(* IEC 61131-3 sources: plc-st-coding-agent/progress/evidence/f14_v11_public_20261113/jobs/custom_deepseek-v4pro (part 2) *)

(* ---- public-hard-02.candidate_03.st ---- *)
TYPE ProcessControl_State : (PC_IDLE, PC_MOVING, PC_WAITING); END_TYPE;

FUNCTION_BLOCK FlexibleProcessingControl
VAR_INPUT
    processLength : USINT;
    sensor1 : BOOL;
    sensor2 : BOOL;
    sensor3 : BOOL;
    sensor4 : BOOL;
    sensor5 : BOOL;
    station1Start : BOOL;
    station2Complete : BOOL;
    station3Complete : BOOL;
    station4Complete : BOOL;
    processSequence : ARRAY[1..8] OF USINT;
END_VAR
VAR_OUTPUT
    conveyorLeft : BOOL;
    conveyorRight : BOOL;
END_VAR
VAR
    state : ProcessControl_State := PC_IDLE;
    currentStation : USINT := 1;
    currentIndex : USINT := 1;
    targetStation : USINT := 0;
    targetSensor : BOOL := FALSE;
    local_rt_start : R_TRIG;
    local_rt_st2 : R_TRIG;
    local_rt_st3 : R_TRIG;
    local_rt_st4 : R_TRIG;
END_VAR

(*
ENGINEERING_CONTRACT
  conveyorLeft / conveyorRight activation: PC_MOVING state and target direction >/< currentStation (PUB001-PUB002).
  Retention/hold: outputs stay on each scan while PC_MOVING until target sensor TRUE (PUB002).
  Explicit reset/deactivation: sensor at target station stops motion and sets both outputs FALSE; next start new product.
  Same-scan priority: start request processed only in PC_IDLE; arrival stop and completion advancement are mutually exclusive by state.
  Units/boundaries: processLength 1..8; processSequence index 1..8; currentStation 1..5; final active entry 5 (PUB003).
  Direction: target > current -> conveyorRight; target < current -> conveyorLeft; target == current -> no movement, treated as arrived.
  Completion edge: rising edge of station2Complete/3/4Complete triggers next step.
  Unspecified: equal consecutive station entries skip movement and wait for completion; simultaneous completion inputs while WAITING use current station only.
*)

(* CONTRACT_RULES [] *)

local_rt_start(CLK := station1Start AND sensor1);
local_rt_st2(CLK := station2Complete);
local_rt_st3(CLK := station3Complete);
local_rt_st4(CLK := station4Complete);

CASE state OF
    PC_IDLE:
        conveyorLeft := FALSE;
        conveyorRight := FALSE;
        IF local_rt_start.Q THEN
            currentIndex := 1;
            currentStation := 1;
            targetStation := processSequence[currentIndex];
            IF targetStation = currentStation THEN
                IF targetStation = 5 THEN
                    state := PC_IDLE;
                ELSE
                    state := PC_WAITING;
                END_IF;
            ELSE
                state := PC_MOVING;
            END_IF;
        END_IF;

    PC_MOVING:
        targetSensor := FALSE;
        CASE targetStation OF
            2: targetSensor := sensor2;
            3: targetSensor := sensor3;
            4: targetSensor := sensor4;
            5: targetSensor := sensor5;
        END_CASE;

        IF targetStation > currentStation THEN
            conveyorLeft := FALSE;
            conveyorRight := TRUE;
        ELSIF targetStation < currentStation THEN
            conveyorLeft := TRUE;
            conveyorRight := FALSE;
        ELSE
            conveyorLeft := FALSE;
            conveyorRight := FALSE;
        END_IF;

        IF targetSensor THEN
            conveyorLeft := FALSE;
            conveyorRight := FALSE;
            currentStation := targetStation;
            IF targetStation = 5 THEN
                state := PC_IDLE;
            ELSE
                state := PC_WAITING;
            END_IF;
        END_IF;

    PC_WAITING:
        conveyorLeft := FALSE;
        conveyorRight := FALSE;
        IF (currentStation = 2 AND local_rt_st2.Q) OR
           (currentStation = 3 AND local_rt_st3.Q) OR
           (currentStation = 4 AND local_rt_st4.Q) THEN
            IF currentIndex < processLength THEN
                currentIndex := currentIndex + 1;
                targetStation := processSequence[currentIndex];
                IF targetStation = currentStation THEN
                    IF targetStation = 5 THEN
                        state := PC_IDLE;
                    ELSE
                        state := PC_WAITING;
                    END_IF;
                ELSE
                    state := PC_MOVING;
                END_IF;
            ELSE
                state := PC_IDLE;
            END_IF;
        END_IF;
END_CASE;

(* Same-scan output update after any state transition *)
IF state = PC_MOVING THEN
    IF targetStation > currentStation THEN
        conveyorLeft := FALSE;
        conveyorRight := TRUE;
    ELSIF targetStation < currentStation THEN
        conveyorLeft := TRUE;
        conveyorRight := FALSE;
    ELSE
        conveyorLeft := FALSE;
        conveyorRight := FALSE;
    END_IF;
ELSE
    conveyorLeft := FALSE;
    conveyorRight := FALSE;
END_IF;

END_FUNCTION_BLOCK

(* ---- public-hard-02.candidate_04.st ---- *)
TYPE ProcessControl_State : (PC_IDLE, PC_MOVING, PC_WAITING); END_TYPE;

FUNCTION_BLOCK FlexibleProcessingControl
VAR_INPUT
    processLength : USINT;
    sensor1 : BOOL;
    sensor2 : BOOL;
    sensor3 : BOOL;
    sensor4 : BOOL;
    sensor5 : BOOL;
    station1Start : BOOL;
    station2Complete : BOOL;
    station3Complete : BOOL;
    station4Complete : BOOL;
    processSequence : ARRAY[1..8] OF USINT;
END_VAR
VAR_OUTPUT
    conveyorLeft : BOOL;
    conveyorRight : BOOL;
END_VAR
VAR
    state : ProcessControl_State := PC_IDLE;
    currentStation : USINT := 1;
    currentIndex : USINT := 1;
    targetStation : USINT := 0;
    targetSensor : BOOL := FALSE;
    local_rt_start : R_TRIG;
    local_rt_st2 : R_TRIG;
    local_rt_st3 : R_TRIG;
    local_rt_st4 : R_TRIG;
END_VAR

(*
ENGINEERING_CONTRACT
  conveyorLeft / conveyorRight activation: PC_MOVING state and target direction >/< currentStation (PUB001-PUB002).
  Retention/hold: outputs stay on each scan while PC_MOVING until target sensor TRUE (PUB002).
  Explicit reset/deactivation: sensor at target station stops motion and sets both outputs FALSE; next start new product.
  Same-scan priority: start request processed only in PC_IDLE; arrival stop and completion advancement are mutually exclusive by state.
  Units/boundaries: processLength 1..8; processSequence index 1..8; currentStation 1..5; final active entry 5 (PUB003).
  Direction: target > current -> conveyorRight; target < current -> conveyorLeft; target == current -> no movement, treated as arrived.
  Completion edge: rising edge of station2Complete/3/4Complete triggers next step.
  Unspecified: equal consecutive station entries skip movement and wait for completion; simultaneous completion inputs while WAITING use current station only.
  Same-scan start with target sensor already active causes immediate arrival handling without starting conveyor.
*)

(* CONTRACT_RULES [] *)

local_rt_start(CLK := station1Start AND sensor1);
local_rt_st2(CLK := station2Complete);
local_rt_st3(CLK := station3Complete);
local_rt_st4(CLK := station4Complete);

CASE state OF
    PC_IDLE:
        conveyorLeft := FALSE;
        conveyorRight := FALSE;
        IF local_rt_start.Q THEN
            currentIndex := 1;
            currentStation := 1;
            targetStation := processSequence[currentIndex];
            IF targetStation = currentStation THEN
                IF targetStation = 5 THEN
                    state := PC_IDLE;
                ELSE
                    state := PC_WAITING;
                END_IF;
            ELSE
                targetSensor := FALSE;
                CASE targetStation OF
                    2: targetSensor := sensor2;
                    3: targetSensor := sensor3;
                    4: targetSensor := sensor4;
                    5: targetSensor := sensor5;
                END_CASE;
                IF targetSensor THEN
                    currentStation := targetStation;
                    IF targetStation = 5 THEN
                        state := PC_IDLE;
                    ELSE
                        state := PC_WAITING;
                    END_IF;
                ELSE
                    state := PC_MOVING;
                END_IF;
            END_IF;
        END_IF;

    PC_MOVING:
        targetSensor := FALSE;
        CASE targetStation OF
            2: targetSensor := sensor2;
            3: targetSensor := sensor3;
            4: targetSensor := sensor4;
            5: targetSensor := sensor5;
        END_CASE;

        IF targetStation > currentStation THEN
            conveyorLeft := FALSE;
            conveyorRight := TRUE;
        ELSIF targetStation < currentStation THEN
            conveyorLeft := TRUE;
            conveyorRight := FALSE;
        ELSE
            conveyorLeft := FALSE;
            conveyorRight := FALSE;
        END_IF;

        IF targetSensor THEN
            conveyorLeft := FALSE;
            conveyorRight := FALSE;
            currentStation := targetStation;
            IF targetStation = 5 THEN
                state := PC_IDLE;
            ELSE
                state := PC_WAITING;
            END_IF;
        END_IF;

    PC_WAITING:
        conveyorLeft := FALSE;
        conveyorRight := FALSE;
        IF (currentStation = 2 AND local_rt_st2.Q) OR
           (currentStation = 3 AND local_rt_st3.Q) OR
           (currentStation = 4 AND local_rt_st4.Q) THEN
            IF currentIndex < processLength THEN
                currentIndex := currentIndex + 1;
                targetStation := processSequence[currentIndex];
                IF targetStation = currentStation THEN
                    IF targetStation = 5 THEN
                        state := PC_IDLE;
                    ELSE
                        state := PC_WAITING;
                    END_IF;
                ELSE
                    state := PC_MOVING;
                END_IF;
            ELSE
                state := PC_IDLE;
            END_IF;
        END_IF;
END_CASE;

(* Same-scan output update after any state transition *)
IF state = PC_MOVING THEN
    IF targetStation > currentStation THEN
        conveyorLeft := FALSE;
        conveyorRight := TRUE;
    ELSIF targetStation < currentStation THEN
        conveyorLeft := TRUE;
        conveyorRight := FALSE;
    ELSE
        conveyorLeft := FALSE;
        conveyorRight := FALSE;
    END_IF;
ELSE
    conveyorLeft := FALSE;
    conveyorRight := FALSE;
END_IF;

END_FUNCTION_BLOCK

(* ---- public-hard-02.raw_candidate_01.st ---- *)
TYPE ProcessControl_State : (PC_IDLE, PC_MOVING, PC_WAITING); END_TYPE

FUNCTION_BLOCK FlexibleProcessingControl
VAR_INPUT
    processLength : USINT;
    sensor1 : BOOL;
    sensor2 : BOOL;
    sensor3 : BOOL;
    sensor4 : BOOL;
    sensor5 : BOOL;
    station1Start : BOOL;
    station2Complete : BOOL;
    station3Complete : BOOL;
    station4Complete : BOOL;
    processSequence : ARRAY[1..8] OF USINT;
END_VAR
VAR_OUTPUT
    conveyorLeft : BOOL;
    conveyorRight : BOOL;
END_VAR
VAR
    state : ProcessControl_State := PC_IDLE;
    currentStation : USINT := 1;
    currentIndex : USINT := 1;
    targetStation : USINT := 0;
    targetSensor : BOOL := FALSE;
    local_rt_start : R_TRIG;
    local_rt_st2 : R_TRIG;
    local_rt_st3 : R_TRIG;
    local_rt_st4 : R_TRIG;
END_VAR

(*
ENGINEERING_CONTRACT
  conveyorLeft / conveyorRight activation: PC_MOVING state and target direction >/< currentStation (PUB001-PUB002).
  Retention/hold: outputs stay on each scan while PC_MOVING until target sensor TRUE (PUB002).
  Explicit reset/deactivation: sensor at target station stops motion and sets both outputs FALSE; next start new product.
  Same-scan priority: start request processed only in PC_IDLE; arrival stop and completion advancement are mutually exclusive by state.
  Units/boundaries: processLength 1..8; processSequence index 1..8; currentStation 1..5; final active entry 5 (PUB003).
  Direction: target > current -> conveyorRight; target < current -> conveyorLeft; target == current -> no movement, treated as arrived.
  Completion edge: rising edge of station2Complete/3/4Complete triggers next step.
  Unspecified: equal consecutive station entries skip movement and wait for completion; simultaneous completion inputs while WAITING use current station only.
*)

(* CONTRACT_RULES [] *)

local_rt_start(CLK := station1Start);
local_rt_st2(CLK := station2Complete);
local_rt_st3(CLK := station3Complete);
local_rt_st4(CLK := station4Complete);

CASE state OF
    PC_IDLE:
        conveyorLeft := FALSE;
        conveyorRight := FALSE;
        IF local_rt_start.Q AND sensor1 THEN
            currentIndex := 1;
            currentStation := 1;
            targetStation := processSequence[currentIndex];
            IF targetStation = currentStation THEN
                IF targetStation = 5 THEN
                    state := PC_IDLE;
                ELSE
                    state := PC_WAITING;
                END_IF;
            ELSE
                state := PC_MOVING;
            END_IF;
        END_IF;

    PC_MOVING:
        targetSensor := FALSE;
        CASE targetStation OF
            2: targetSensor := sensor2;
            3: targetSensor := sensor3;
            4: targetSensor := sensor4;
            5: targetSensor := sensor5;
        END_CASE;

        IF targetStation > currentStation THEN
            conveyorLeft := FALSE;
            conveyorRight := TRUE;
        ELSIF targetStation < currentStation THEN
            conveyorLeft := TRUE;
            conveyorRight := FALSE;
        ELSE
            conveyorLeft := FALSE;
            conveyorRight := FALSE;
        END_IF;

        IF targetSensor THEN
            conveyorLeft := FALSE;
            conveyorRight := FALSE;
            currentStation := targetStation;
            IF targetStation = 5 THEN
                state := PC_IDLE;
            ELSE
                state := PC_WAITING;
            END_IF;
        END_IF;

    PC_WAITING:
        conveyorLeft := FALSE;
        conveyorRight := FALSE;
        IF (currentStation = 2 AND local_rt_st2.Q) OR
           (currentStation = 3 AND local_rt_st3.Q) OR
           (currentStation = 4 AND local_rt_st4.Q) THEN
            IF currentIndex < processLength THEN
                currentIndex := currentIndex + 1;
                targetStation := processSequence[currentIndex];
                IF targetStation = currentStation THEN
                    IF targetStation = 5 THEN
                        state := PC_IDLE;
                    ELSE
                        state := PC_WAITING;
                    END_IF;
                ELSE
                    state := PC_MOVING;
                END_IF;
            ELSE
                state := PC_IDLE;
            END_IF;
        END_IF;
END_CASE;

(* ---- public-hard-02.raw_candidate_02.st ---- *)
TYPE ProcessControl_State : (PC_IDLE, PC_MOVING, PC_WAITING); END_TYPE;

FUNCTION_BLOCK FlexibleProcessingControl
VAR_INPUT
    processLength : USINT;
    sensor1 : BOOL;
    sensor2 : BOOL;
    sensor3 : BOOL;
    sensor4 : BOOL;
    sensor5 : BOOL;
    station1Start : BOOL;
    station2Complete : BOOL;
    station3Complete : BOOL;
    station4Complete : BOOL;
    processSequence : ARRAY[1..8] OF USINT;
END_VAR
VAR_OUTPUT
    conveyorLeft : BOOL;
    conveyorRight : BOOL;
END_VAR
VAR
    state : ProcessControl_State := PC_IDLE;
    currentStation : USINT := 1;
    currentIndex : USINT := 1;
    targetStation : USINT := 0;
    targetSensor : BOOL := FALSE;
    local_rt_start : R_TRIG;
    local_rt_st2 : R_TRIG;
    local_rt_st3 : R_TRIG;
    local_rt_st4 : R_TRIG;
END_VAR

(*
ENGINEERING_CONTRACT
  conveyorLeft / conveyorRight activation: PC_MOVING state and target direction >/< currentStation (PUB001-PUB002).
  Retention/hold: outputs stay on each scan while PC_MOVING until target sensor TRUE (PUB002).
  Explicit reset/deactivation: sensor at target station stops motion and sets both outputs FALSE; next start new product.
  Same-scan priority: start request processed only in PC_IDLE; arrival stop and completion advancement are mutually exclusive by state.
  Units/boundaries: processLength 1..8; processSequence index 1..8; currentStation 1..5; final active entry 5 (PUB003).
  Direction: target > current -> conveyorRight; target < current -> conveyorLeft; target == current -> no movement, treated as arrived.
  Completion edge: rising edge of station2Complete/3/4Complete triggers next step.
  Unspecified: equal consecutive station entries skip movement and wait for completion; simultaneous completion inputs while WAITING use current station only.
*)

(* CONTRACT_RULES [] *)

local_rt_start(CLK := station1Start);
local_rt_st2(CLK := station2Complete);
local_rt_st3(CLK := station3Complete);
local_rt_st4(CLK := station4Complete);

CASE state OF
    PC_IDLE:
        conveyorLeft := FALSE;
        conveyorRight := FALSE;
        IF local_rt_start.Q AND sensor1 THEN
            currentIndex := 1;
            currentStation := 1;
            targetStation := processSequence[currentIndex];
            IF targetStation = currentStation THEN
                IF targetStation = 5 THEN
                    state := PC_IDLE;
                ELSE
                    state := PC_WAITING;
                END_IF;
            ELSE
                state := PC_MOVING;
            END_IF;
        END_IF;

    PC_MOVING:
        targetSensor := FALSE;
        CASE targetStation OF
            2: targetSensor := sensor2;
            3: targetSensor := sensor3;
            4: targetSensor := sensor4;
            5: targetSensor := sensor5;
        END_CASE;

        IF targetStation > currentStation THEN
            conveyorLeft := FALSE;
            conveyorRight := TRUE;
        ELSIF targetStation < currentStation THEN
            conveyorLeft := TRUE;
            conveyorRight := FALSE;
        ELSE
            conveyorLeft := FALSE;
            conveyorRight := FALSE;
        END_IF;

        IF targetSensor THEN
            conveyorLeft := FALSE;
            conveyorRight := FALSE;
            currentStation := targetStation;
            IF targetStation = 5 THEN
                state := PC_IDLE;
            ELSE
                state := PC_WAITING;
            END_IF;
        END_IF;

    PC_WAITING:
        conveyorLeft := FALSE;
        conveyorRight := FALSE;
        IF (currentStation = 2 AND local_rt_st2.Q) OR
           (currentStation = 3 AND local_rt_st3.Q) OR
           (currentStation = 4 AND local_rt_st4.Q) THEN
            IF currentIndex < processLength THEN
                currentIndex := currentIndex + 1;
                targetStation := processSequence[currentIndex];
                IF targetStation = currentStation THEN
                    IF targetStation = 5 THEN
                        state := PC_IDLE;
                    ELSE
                        state := PC_WAITING;
                    END_IF;
                ELSE
                    state := PC_MOVING;
                END_IF;
            ELSE
                state := PC_IDLE;
            END_IF;
        END_IF;
END_CASE;

END_FUNCTION_BLOCK

(* ---- public-hard-02.raw_candidate_03.st ---- *)
TYPE ProcessControl_State : (PC_IDLE, PC_MOVING, PC_WAITING); END_TYPE;

FUNCTION_BLOCK FlexibleProcessingControl
VAR_INPUT
    processLength : USINT;
    sensor1 : BOOL;
    sensor2 : BOOL;
    sensor3 : BOOL;
    sensor4 : BOOL;
    sensor5 : BOOL;
    station1Start : BOOL;
    station2Complete : BOOL;
    station3Complete : BOOL;
    station4Complete : BOOL;
    processSequence : ARRAY[1..8] OF USINT;
END_VAR
VAR_OUTPUT
    conveyorLeft : BOOL;
    conveyorRight : BOOL;
END_VAR
VAR
    state : ProcessControl_State := PC_IDLE;
    currentStation : USINT := 1;
    currentIndex : USINT := 1;
    targetStation : USINT := 0;
    targetSensor : BOOL := FALSE;
    local_rt_start : R_TRIG;
    local_rt_st2 : R_TRIG;
    local_rt_st3 : R_TRIG;
    local_rt_st4 : R_TRIG;
END_VAR

(*
ENGINEERING_CONTRACT
  conveyorLeft / conveyorRight activation: PC_MOVING state and target direction >/< currentStation (PUB001-PUB002).
  Retention/hold: outputs stay on each scan while PC_MOVING until target sensor TRUE (PUB002).
  Explicit reset/deactivation: sensor at target station stops motion and sets both outputs FALSE; next start new product.
  Same-scan priority: start request processed only in PC_IDLE; arrival stop and completion advancement are mutually exclusive by state.
  Units/boundaries: processLength 1..8; processSequence index 1..8; currentStation 1..5; final active entry 5 (PUB003).
  Direction: target > current -> conveyorRight; target < current -> conveyorLeft; target == current -> no movement, treated as arrived.
  Completion edge: rising edge of station2Complete/3/4Complete triggers next step.
  Unspecified: equal consecutive station entries skip movement and wait for completion; simultaneous completion inputs while WAITING use current station only.
*)

(* CONTRACT_RULES [] *)

local_rt_start(CLK := station1Start AND sensor1);
local_rt_st2(CLK := station2Complete);
local_rt_st3(CLK := station3Complete);
local_rt_st4(CLK := station4Complete);

CASE state OF
    PC_IDLE:
        conveyorLeft := FALSE;
        conveyorRight := FALSE;
        IF local_rt_start.Q THEN
            currentIndex := 1;
            currentStation := 1;
            targetStation := processSequence[currentIndex];
            IF targetStation = currentStation THEN
                IF targetStation = 5 THEN
                    state := PC_IDLE;
                ELSE
                    state := PC_WAITING;
                END_IF;
            ELSE
                state := PC_MOVING;
            END_IF;
        END_IF;

    PC_MOVING:
        targetSensor := FALSE;
        CASE targetStation OF
            2: targetSensor := sensor2;
            3: targetSensor := sensor3;
            4: targetSensor := sensor4;
            5: targetSensor := sensor5;
        END_CASE;

        IF targetStation > currentStation THEN
            conveyorLeft := FALSE;
            conveyorRight := TRUE;
        ELSIF targetStation < currentStation THEN
            conveyorLeft := TRUE;
            conveyorRight := FALSE;
        ELSE
            conveyorLeft := FALSE;
            conveyorRight := FALSE;
        END_IF;

        IF targetSensor THEN
            conveyorLeft := FALSE;
            conveyorRight := FALSE;
            currentStation := targetStation;
            IF targetStation = 5 THEN
                state := PC_IDLE;
            ELSE
                state := PC_WAITING;
            END_IF;
        END_IF;

    PC_WAITING:
        conveyorLeft := FALSE;
        conveyorRight := FALSE;
        IF (currentStation = 2 AND local_rt_st2.Q) OR
           (currentStation = 3 AND local_rt_st3.Q) OR
           (currentStation = 4 AND local_rt_st4.Q) THEN
            IF currentIndex < processLength THEN
                currentIndex := currentIndex + 1;
                targetStation := processSequence[currentIndex];
                IF targetStation = currentStation THEN
                    IF targetStation = 5 THEN
                        state := PC_IDLE;
                    ELSE
                        state := PC_WAITING;
                    END_IF;
                ELSE
                    state := PC_MOVING;
                END_IF;
            ELSE
                state := PC_IDLE;
            END_IF;
        END_IF;
END_CASE;

(* Same-scan output update after any state transition *)
IF state = PC_MOVING THEN
    IF targetStation > currentStation THEN
        conveyorLeft := FALSE;
        conveyorRight := TRUE;
    ELSIF targetStation < currentStation THEN
        conveyorLeft := TRUE;
        conveyorRight := FALSE;
    ELSE
        conveyorLeft := FALSE;
        conveyorRight := FALSE;
    END_IF;
ELSE
    conveyorLeft := FALSE;
    conveyorRight := FALSE;
END_IF;

END_FUNCTION_BLOCK

(* ---- public-hard-02.raw_candidate_04.st ---- *)
TYPE ProcessControl_State : (PC_IDLE, PC_MOVING, PC_WAITING); END_TYPE;

FUNCTION_BLOCK FlexibleProcessingControl
VAR_INPUT
    processLength : USINT;
    sensor1 : BOOL;
    sensor2 : BOOL;
    sensor3 : BOOL;
    sensor4 : BOOL;
    sensor5 : BOOL;
    station1Start : BOOL;
    station2Complete : BOOL;
    station3Complete : BOOL;
    station4Complete : BOOL;
    processSequence : ARRAY[1..8] OF USINT;
END_VAR
VAR_OUTPUT
    conveyorLeft : BOOL;
    conveyorRight : BOOL;
END_VAR
VAR
    state : ProcessControl_State := PC_IDLE;
    currentStation : USINT := 1;
    currentIndex : USINT := 1;
    targetStation : USINT := 0;
    targetSensor : BOOL := FALSE;
    local_rt_start : R_TRIG;
    local_rt_st2 : R_TRIG;
    local_rt_st3 : R_TRIG;
    local_rt_st4 : R_TRIG;
END_VAR

(*
ENGINEERING_CONTRACT
  conveyorLeft / conveyorRight activation: PC_MOVING state and target direction >/< currentStation (PUB001-PUB002).
  Retention/hold: outputs stay on each scan while PC_MOVING until target sensor TRUE (PUB002).
  Explicit reset/deactivation: sensor at target station stops motion and sets both outputs FALSE; next start new product.
  Same-scan priority: start request processed only in PC_IDLE; arrival stop and completion advancement are mutually exclusive by state.
  Units/boundaries: processLength 1..8; processSequence index 1..8; currentStation 1..5; final active entry 5 (PUB003).
  Direction: target > current -> conveyorRight; target < current -> conveyorLeft; target == current -> no movement, treated as arrived.
  Completion edge: rising edge of station2Complete/3/4Complete triggers next step.
  Unspecified: equal consecutive station entries skip movement and wait for completion; simultaneous completion inputs while WAITING use current station only.
  Same-scan start with target sensor already active causes immediate arrival handling without starting conveyor.
*)

(* CONTRACT_RULES [] *)

local_rt_start(CLK := station1Start AND sensor1);
local_rt_st2(CLK := station2Complete);
local_rt_st3(CLK := station3Complete);
local_rt_st4(CLK := station4Complete);

CASE state OF
    PC_IDLE:
        conveyorLeft := FALSE;
        conveyorRight := FALSE;
        IF local_rt_start.Q THEN
            currentIndex := 1;
            currentStation := 1;
            targetStation := processSequence[currentIndex];
            IF targetStation = currentStation THEN
                IF targetStation = 5 THEN
                    state := PC_IDLE;
                ELSE
                    state := PC_WAITING;
                END_IF;
            ELSE
                targetSensor := FALSE;
                CASE targetStation OF
                    2: targetSensor := sensor2;
                    3: targetSensor := sensor3;
                    4: targetSensor := sensor4;
                    5: targetSensor := sensor5;
                END_CASE;
                IF targetSensor THEN
                    currentStation := targetStation;
                    IF targetStation = 5 THEN
                        state := PC_IDLE;
                    ELSE
                        state := PC_WAITING;
                    END_IF;
                ELSE
                    state := PC_MOVING;
                END_IF;
            END_IF;
        END_IF;

    PC_MOVING:
        targetSensor := FALSE;
        CASE targetStation OF
            2: targetSensor := sensor2;
            3: targetSensor := sensor3;
            4: targetSensor := sensor4;
            5: targetSensor := sensor5;
        END_CASE;

        IF targetStation > currentStation THEN
            conveyorLeft := FALSE;
            conveyorRight := TRUE;
        ELSIF targetStation < currentStation THEN
            conveyorLeft := TRUE;
            conveyorRight := FALSE;
        ELSE
            conveyorLeft := FALSE;
            conveyorRight := FALSE;
        END_IF;

        IF targetSensor THEN
            conveyorLeft := FALSE;
            conveyorRight := FALSE;
            currentStation := targetStation;
            IF targetStation = 5 THEN
                state := PC_IDLE;
            ELSE
                state := PC_WAITING;
            END_IF;
        END_IF;

    PC_WAITING:
        conveyorLeft := FALSE;
        conveyorRight := FALSE;
        IF (currentStation = 2 AND local_rt_st2.Q) OR
           (currentStation = 3 AND local_rt_st3.Q) OR
           (currentStation = 4 AND local_rt_st4.Q) THEN
            IF currentIndex < processLength THEN
                currentIndex := currentIndex + 1;
                targetStation := processSequence[currentIndex];
                IF targetStation = currentStation THEN
                    IF targetStation = 5 THEN
                        state := PC_IDLE;
                    ELSE
                        state := PC_WAITING;
                    END_IF;
                ELSE
                    state := PC_MOVING;
                END_IF;
            ELSE
                state := PC_IDLE;
            END_IF;
        END_IF;
END_CASE;

(* Same-scan output update after any state transition *)
IF state = PC_MOVING THEN
    IF targetStation > currentStation THEN
        conveyorLeft := FALSE;
        conveyorRight := TRUE;
    ELSIF targetStation < currentStation THEN
        conveyorLeft := TRUE;
        conveyorRight := FALSE;
    ELSE
        conveyorLeft := FALSE;
        conveyorRight := FALSE;
    END_IF;
ELSE
    conveyorLeft := FALSE;
    conveyorRight := FALSE;
END_IF;

END_FUNCTION_BLOCK

(* ---- public-hard-03.candidate_01.st ---- *)
TYPE ST_Recipe :
STRUCT
    recipeID : INT;
    ingredientType : INT;
    ingredientRatio : REAL;
    productionTemperature : REAL;
END_STRUCT
END_TYPE;

FUNCTION_BLOCK RecipeManagement
VAR_INPUT
    addRecipe : BOOL;
    deleteRecipe : BOOL;
    modifyRecipe : BOOL;
    queryRecipe : BOOL;
    recipeIn : ST_Recipe;
END_VAR
VAR_OUTPUT
    recipeAdded : BOOL;
    recipeDeleted : BOOL;
    recipeModified : BOOL;
    recipeQueryResult : ST_Recipe;
    error : BOOL;
    status : WORD;
END_VAR
VAR_IN_OUT
    recipe : ARRAY[1..10] OF ST_Recipe;
END_VAR
VAR
    tmp_i : INT;
    tmp_idx : INT;
    tmp_empty : INT;
    tmp_duplicate : BOOL;
    tmp_count : INT;
END_VAR

(* ENGINEERING_CONTRACT
   Pub outputs recipeAdded/Deleted/Modified are one-scan success pulses; no latch.
   error/status are combinational: FALSE/0 on success or idle, TRUE/code on specified failure.
   recipe array persists in IN_OUT slots. Add uses first empty slot; delete clears ID only; modify replaces whole recipe.
   Query/delete/modify search only non-zero recipeID; add duplicate check includes recipeID 0 as empty-slot duplicate.
   Multiple simultaneous request inputs are unspecified; implementation reports error=TRUE, status=16#8000 and performs none.
   Boundary: recipeID 0 is never a queryable/deletable/modifiable identifier.
*)
(* CONTRACT_RULES [] *)

recipeAdded := FALSE;
recipeDeleted := FALSE;
recipeModified := FALSE;
error := FALSE;
status := 0;
recipeQueryResult.recipeID := 0;
recipeQueryResult.ingredientType := 0;
recipeQueryResult.ingredientRatio := 0.0;
recipeQueryResult.productionTemperature := 0.0;

tmp_count := 0;
IF addRecipe THEN
    tmp_count := tmp_count + 1;
END_IF;
IF deleteRecipe THEN
    tmp_count := tmp_count + 1;
END_IF;
IF modifyRecipe THEN
    tmp_count := tmp_count + 1;
END_IF;
IF queryRecipe THEN
    tmp_count := tmp_count + 1;
END_IF;

IF tmp_count > 1 THEN
    error := TRUE;
    status := 16#8000;
    RETURN;
END_IF;

IF addRecipe THEN
    tmp_duplicate := FALSE;
    FOR tmp_i := 1 TO 10 DO
        IF recipe[tmp_i].recipeID = recipeIn.recipeID THEN
            tmp_duplicate := TRUE;
            EXIT;
        END_IF;
    END_FOR;

    IF tmp_duplicate THEN
        error := TRUE;
        status := 16#8002;
    ELSE
        tmp_empty := 0;
        FOR tmp_i := 1 TO 10 DO
            IF recipe[tmp_i].recipeID = 0 THEN
                tmp_empty := tmp_i;
                EXIT;
            END_IF;
        END_FOR;

        IF tmp_empty = 0 THEN
            error := TRUE;
            status := 16#8003;
        ELSE
            recipe[tmp_empty] := recipeIn;
            recipeAdded := TRUE;
        END_IF;
    END_IF;

ELSIF deleteRecipe THEN
    tmp_idx := 0;
    IF recipeIn.recipeID <> 0 THEN
        FOR tmp_i := 1 TO 10 DO
            IF recipe[tmp_i].recipeID = recipeIn.recipeID THEN
                tmp_idx := tmp_i;
                EXIT;
            END_IF;
        END_FOR;
    END_IF;

    IF tmp_idx = 0 THEN
        error := TRUE;
        status := 16#8004;
    ELSE
        recipe[tmp_idx].recipeID := 0;
        recipeDeleted := TRUE;
    END_IF;

ELSIF modifyRecipe THEN
    tmp_idx := 0;
    IF recipeIn.recipeID <> 0 THEN
        FOR tmp_i := 1 TO 10 DO
            IF recipe[tmp_i].recipeID = recipeIn.recipeID THEN
                tmp_idx := tmp_i;
                EXIT;
            END_IF;
        END_FOR;
    END_IF;

    IF tmp_idx = 0 THEN
        error := TRUE;
        status := 16#8005;
    ELSE
        recipe[tmp_idx] := recipeIn;
        recipeModified := TRUE;
    END_IF;

ELSIF queryRecipe THEN
    tmp_idx := 0;
    IF recipeIn.recipeID <> 0 THEN
        FOR tmp_i := 1 TO 10 DO
            IF recipe[tmp_i].recipeID = recipeIn.recipeID THEN
                tmp_idx := tmp_i;
                EXIT;
            END_IF;
        END_FOR;
    END_IF;

    IF tmp_idx = 0 THEN
        error := TRUE;
        status := 16#8001;
    ELSE
        recipeQueryResult := recipe[tmp_idx];
    END_IF;
END_IF;

(* ---- public-hard-03.candidate_02.st ---- *)
TYPE ST_Recipe :
STRUCT
    recipeID : INT;
    ingredientType : INT;
    ingredientRatio : REAL;
    productionTemperature : REAL;
END_STRUCT
END_TYPE;

FUNCTION_BLOCK RecipeManagement
VAR_INPUT
    addRecipe : BOOL;
    deleteRecipe : BOOL;
    modifyRecipe : BOOL;
    queryRecipe : BOOL;
    recipeIn : ST_Recipe;
END_VAR
VAR_OUTPUT
    recipeAdded : BOOL;
    recipeDeleted : BOOL;
    recipeModified : BOOL;
    recipeQueryResult : ST_Recipe;
    error : BOOL;
    status : WORD;
END_VAR
VAR_IN_OUT
    recipe : ARRAY[1..10] OF ST_Recipe;
END_VAR
VAR
    tmp_i : INT;
    tmp_idx : INT;
    tmp_empty : INT;
    tmp_duplicate : BOOL;
    tmp_count : INT;
END_VAR

(* ENGINEERING_CONTRACT
   Pub outputs recipeAdded/Deleted/Modified are one-scan success pulses; no latch.
   error/status are combinational: FALSE/0 on success or idle, TRUE/code on specified failure.
   recipe array persists in IN_OUT slots. Add uses first empty slot; delete clears ID only; modify replaces whole recipe.
   Query/delete/modify search only non-zero recipeID; add duplicate check includes recipeID 0 as empty-slot duplicate.
   Multiple simultaneous request inputs are unspecified; implementation reports error=TRUE, status=16#8000 and performs none.
   Boundary: recipeID 0 is never a queryable/deletable/modifiable identifier.
*)
(* CONTRACT_RULES [] *)

recipeAdded := FALSE;
recipeDeleted := FALSE;
recipeModified := FALSE;
error := FALSE;
status := 0;
recipeQueryResult.recipeID := 0;
recipeQueryResult.ingredientType := 0;
recipeQueryResult.ingredientRatio := 0.0;
recipeQueryResult.productionTemperature := 0.0;

tmp_count := 0;
IF addRecipe THEN
    tmp_count := tmp_count + 1;
END_IF;
IF deleteRecipe THEN
    tmp_count := tmp_count + 1;
END_IF;
IF modifyRecipe THEN
    tmp_count := tmp_count + 1;
END_IF;
IF queryRecipe THEN
    tmp_count := tmp_count + 1;
END_IF;

IF tmp_count > 1 THEN
    error := TRUE;
    status := 16#8000;
    RETURN;
END_IF;

IF addRecipe THEN
    tmp_duplicate := FALSE;
    FOR tmp_i := 1 TO 10 DO
        IF recipe[tmp_i].recipeID = recipeIn.recipeID THEN
            tmp_duplicate := TRUE;
            EXIT;
        END_IF;
    END_FOR;

    IF tmp_duplicate THEN
        error := TRUE;
        status := 16#8002;
    ELSE
        tmp_empty := 0;
        FOR tmp_i := 1 TO 10 DO
            IF recipe[tmp_i].recipeID = 0 THEN
                tmp_empty := tmp_i;
                EXIT;
            END_IF;
        END_FOR;

        IF tmp_empty = 0 THEN
            error := TRUE;
            status := 16#8003;
        ELSE
            recipe[tmp_empty] := recipeIn;
            recipeAdded := TRUE;
        END_IF;
    END_IF;

ELSIF deleteRecipe THEN
    tmp_idx := 0;
    IF recipeIn.recipeID <> 0 THEN
        FOR tmp_i := 1 TO 10 DO
            IF recipe[tmp_i].recipeID = recipeIn.recipeID THEN
                tmp_idx := tmp_i;
                EXIT;
            END_IF;
        END_FOR;
    END_IF;

    IF tmp_idx = 0 THEN
        error := TRUE;
        status := 16#8004;
    ELSE
        recipe[tmp_idx].recipeID := 0;
        recipeDeleted := TRUE;
    END_IF;

ELSIF modifyRecipe THEN
    tmp_idx := 0;
    IF recipeIn.recipeID <> 0 THEN
        FOR tmp_i := 1 TO 10 DO
            IF recipe[tmp_i].recipeID = recipeIn.recipeID THEN
                tmp_idx := tmp_i;
                EXIT;
            END_IF;
        END_FOR;
    END_IF;

    IF tmp_idx = 0 THEN
        error := TRUE;
        status := 16#8005;
    ELSE
        recipe[tmp_idx] := recipeIn;
        recipeModified := TRUE;
    END_IF;

ELSIF queryRecipe THEN
    tmp_idx := 0;
    IF recipeIn.recipeID <> 0 THEN
        FOR tmp_i := 1 TO 10 DO
            IF recipe[tmp_i].recipeID = recipeIn.recipeID THEN
                tmp_idx := tmp_i;
                EXIT;
            END_IF;
        END_FOR;
    END_IF;

    IF tmp_idx = 0 THEN
        error := TRUE;
        status := 16#8001;
    ELSE
        recipeQueryResult := recipe[tmp_idx];
    END_IF;
END_IF;

END_FUNCTION_BLOCK

(* ---- public-hard-03.candidate_03.st ---- *)
TYPE ST_Recipe :
STRUCT
    recipeID : INT;
    ingredientType : INT;
    ingredientRatio : REAL;
    productionTemperature : REAL;
END_STRUCT
END_TYPE;

FUNCTION_BLOCK RecipeManagement
VAR_INPUT
    addRecipe : BOOL;
    deleteRecipe : BOOL;
    modifyRecipe : BOOL;
    queryRecipe : BOOL;
    recipeIn : ST_Recipe;
END_VAR
VAR_OUTPUT
    recipeAdded : BOOL;
    recipeDeleted : BOOL;
    recipeModified : BOOL;
    recipeQueryResult : ST_Recipe;
    error : BOOL;
    status : WORD;
END_VAR
VAR_IN_OUT
    recipe : ARRAY[1..10] OF ST_Recipe;
END_VAR
VAR
    trg_add : R_TRIG;
    trg_delete : R_TRIG;
    trg_modify : R_TRIG;
    trg_query : R_TRIG;
    tmp_i : INT;
    tmp_idx : INT;
    tmp_empty : INT;
    tmp_duplicate : BOOL;
    tmp_count : INT;
END_VAR

(* ENGINEERING_CONTRACT
   Pub outputs recipeAdded/Deleted/Modified are one-scan success pulses; no latch.
   error/status are combinational: FALSE/0 on success or idle, TRUE/code on specified failure.
   recipe array persists in IN_OUT slots. Add uses first empty slot; delete clears ID only; modify replaces whole recipe.
   Query/delete/modify search only non-zero recipeID; add duplicate check includes recipeID 0 as empty-slot duplicate.
   Multiple simultaneous request inputs are unspecified; implementation reports error=TRUE, status=16#8000 and performs none.
   Boundary: recipeID 0 is never a queryable/deletable/modifiable identifier.
*)
(* CONTRACT_RULES [] *)

trg_add(CLK := addRecipe);
trg_delete(CLK := deleteRecipe);
trg_modify(CLK := modifyRecipe);
trg_query(CLK := queryRecipe);

recipeAdded := FALSE;
recipeDeleted := FALSE;
recipeModified := FALSE;
error := FALSE;
status := 0;
recipeQueryResult.recipeID := 0;
recipeQueryResult.ingredientType := 0;
recipeQueryResult.ingredientRatio := 0.0;
recipeQueryResult.productionTemperature := 0.0;

tmp_count := 0;
IF trg_add.Q THEN
    tmp_count := tmp_count + 1;
END_IF;
IF trg_delete.Q THEN
    tmp_count := tmp_count + 1;
END_IF;
IF trg_modify.Q THEN
    tmp_count := tmp_count + 1;
END_IF;
IF trg_query.Q THEN
    tmp_count := tmp_count + 1;
END_IF;

IF tmp_count > 1 THEN
    error := TRUE;
    status := 16#8000;
    RETURN;
END_IF;

IF trg_add.Q THEN
    tmp_duplicate := FALSE;
    FOR tmp_i := 1 TO 10 DO
        IF recipe[tmp_i].recipeID = recipeIn.recipeID THEN
            tmp_duplicate := TRUE;
            EXIT;
        END_IF;
    END_FOR;

    IF tmp_duplicate THEN
        error := TRUE;
        status := 16#8002;
    ELSE
        tmp_empty := 0;
        FOR tmp_i := 1 TO 10 DO
            IF recipe[tmp_i].recipeID = 0 THEN
                tmp_empty := tmp_i;
                EXIT;
            END_IF;
        END_FOR;

        IF tmp_empty = 0 THEN
            error := TRUE;
            status := 16#8003;
        ELSE
            recipe[tmp_empty] := recipeIn;
            recipeAdded := TRUE;
        END_IF;
    END_IF;

ELSIF trg_delete.Q THEN
    tmp_idx := 0;
    IF recipeIn.recipeID <> 0 THEN
        FOR tmp_i := 1 TO 10 DO
            IF recipe[tmp_i].recipeID = recipeIn.recipeID THEN
                tmp_idx := tmp_i;
                EXIT;
            END_IF;
        END_FOR;
    END_IF;

    IF tmp_idx = 0 THEN
        error := TRUE;
        status := 16#8004;
    ELSE
        recipe[tmp_idx].recipeID := 0;
        recipeDeleted := TRUE;
    END_IF;

ELSIF trg_modify.Q THEN
    tmp_idx := 0;
    IF recipeIn.recipeID <> 0 THEN
        FOR tmp_i := 1 TO 10 DO
            IF recipe[tmp_i].recipeID = recipeIn.recipeID THEN
                tmp_idx := tmp_i;
                EXIT;
            END_IF;
        END_FOR;
    END_IF;

    IF tmp_idx = 0 THEN
        error := TRUE;
        status := 16#8005;
    ELSE
        recipe[tmp_idx] := recipeIn;
        recipeModified := TRUE;
    END_IF;

ELSIF trg_query.Q THEN
    tmp_idx := 0;
    IF recipeIn.recipeID <> 0 THEN
        FOR tmp_i := 1 TO 10 DO
            IF recipe[tmp_i].recipeID = recipeIn.recipeID THEN
                tmp_idx := tmp_i;
                EXIT;
            END_IF;
        END_FOR;
    END_IF;

    IF tmp_idx = 0 THEN
        error := TRUE;
        status := 16#8001;
    ELSE
        recipeQueryResult := recipe[tmp_idx];
    END_IF;
END_IF;

END_FUNCTION_BLOCK

(* ---- public-hard-03.candidate_04.st ---- *)
TYPE ST_Recipe :
STRUCT
    recipeID : INT;
    ingredientType : INT;
    ingredientRatio : REAL;
    productionTemperature : REAL;
END_STRUCT
END_TYPE;

FUNCTION_BLOCK RecipeManagement
VAR_INPUT
    addRecipe : BOOL;
    deleteRecipe : BOOL;
    modifyRecipe : BOOL;
    queryRecipe : BOOL;
    recipeIn : ST_Recipe;
END_VAR
VAR_OUTPUT
    recipeAdded : BOOL;
    recipeDeleted : BOOL;
    recipeModified : BOOL;
    recipeQueryResult : ST_Recipe;
    error : BOOL;
    status : WORD;
END_VAR
VAR_IN_OUT
    recipe : ARRAY[1..10] OF ST_Recipe;
END_VAR
VAR
    trg_add : R_TRIG;
    trg_delete : R_TRIG;
    trg_modify : R_TRIG;
    trg_query : R_TRIG;
    tmp_i : INT;
    tmp_idx : INT;
    tmp_empty : INT;
    tmp_duplicate : BOOL;
    tmp_count : INT;
END_VAR

(* ENGINEERING_CONTRACT
   Pub outputs recipeAdded/Deleted/Modified are one-scan success pulses; no latch.
   error/status are combinational: FALSE/0 on success or idle, TRUE/code on specified failure.
   recipe array persists in IN_OUT slots. Add uses first empty slot; delete clears ID only; modify replaces whole recipe.
   Query/delete/modify search only non-zero recipeID; add duplicate check includes recipeID 0 as empty-slot duplicate.
   Multiple simultaneous request inputs are unspecified; implementation reports error=TRUE, status=16#8000 and performs none.
   Boundary: recipeID 0 is never a queryable/deletable/modifiable identifier.
   recipeQueryResult is retained after a successful query until the next successful query. It is not cleared on idle or on an unsuccessful query.
*)
(* CONTRACT_RULES [] *)

trg_add(CLK := addRecipe);
trg_delete(CLK := deleteRecipe);
trg_modify(CLK := modifyRecipe);
trg_query(CLK := queryRecipe);

recipeAdded := FALSE;
recipeDeleted := FALSE;
recipeModified := FALSE;
error := FALSE;
status := 0;

tmp_count := 0;
IF trg_add.Q THEN
    tmp_count := tmp_count + 1;
END_IF;
IF trg_delete.Q THEN
    tmp_count := tmp_count + 1;
END_IF;
IF trg_modify.Q THEN
    tmp_count := tmp_count + 1;
END_IF;
IF trg_query.Q THEN
    tmp_count := tmp_count + 1;
END_IF;

IF tmp_count > 1 THEN
    error := TRUE;
    status := 16#8000;
    RETURN;
END_IF;

IF trg_add.Q THEN
    tmp_duplicate := FALSE;
    FOR tmp_i := 1 TO 10 DO
        IF recipe[tmp_i].recipeID = recipeIn.recipeID THEN
            tmp_duplicate := TRUE;
            EXIT;
        END_IF;
    END_FOR;

    IF tmp_duplicate THEN
        error := TRUE;
        status := 16#8002;
    ELSE
        tmp_empty := 0;
        FOR tmp_i := 1 TO 10 DO
            IF recipe[tmp_i].recipeID = 0 THEN
                tmp_empty := tmp_i;
                EXIT;
            END_IF;
        END_FOR;

        IF tmp_empty = 0 THEN
            error := TRUE;
            status := 16#8003;
        ELSE
            recipe[tmp_empty] := recipeIn;
            recipeAdded := TRUE;
        END_IF;
    END_IF;

ELSIF trg_delete.Q THEN
    tmp_idx := 0;
    IF recipeIn.recipeID <> 0 THEN
        FOR tmp_i := 1 TO 10 DO
            IF recipe[tmp_i].recipeID = recipeIn.recipeID THEN
                tmp_idx := tmp_i;
                EXIT;
            END_IF;
        END_FOR;
    END_IF;

    IF tmp_idx = 0 THEN
        error := TRUE;
        status := 16#8004;
    ELSE
        recipe[tmp_idx].recipeID := 0;
        recipeDeleted := TRUE;
    END_IF;

ELSIF trg_modify.Q THEN
    tmp_idx := 0;
    IF recipeIn.recipeID <> 0 THEN
        FOR tmp_i := 1 TO 10 DO
            IF recipe[tmp_i].recipeID = recipeIn.recipeID THEN
                tmp_idx := tmp_i;
                EXIT;
            END_IF;
        END_FOR;
    END_IF;

    IF tmp_idx = 0 THEN
        error := TRUE;
        status := 16#8005;
    ELSE
        recipe[tmp_idx] := recipeIn;
        recipeModified := TRUE;
    END_IF;

ELSIF trg_query.Q THEN
    tmp_idx := 0;
    IF recipeIn.recipeID <> 0 THEN
        FOR tmp_i := 1 TO 10 DO
            IF recipe[tmp_i].recipeID = recipeIn.recipeID THEN
                tmp_idx := tmp_i;
                EXIT;
            END_IF;
        END_FOR;
    END_IF;

    IF tmp_idx = 0 THEN
        error := TRUE;
        status := 16#8001;
    ELSE
        recipeQueryResult := recipe[tmp_idx];
    END_IF;
END_IF;

END_FUNCTION_BLOCK

(* ---- public-hard-03.raw_candidate_01.st ---- *)
TYPE ST_Recipe :
STRUCT
    recipeID : INT;
    ingredientType : INT;
    ingredientRatio : REAL;
    productionTemperature : REAL;
END_STRUCT
END_TYPE

FUNCTION_BLOCK RecipeManagement
VAR_INPUT
    addRecipe : BOOL;
    deleteRecipe : BOOL;
    modifyRecipe : BOOL;
    queryRecipe : BOOL;
    recipeIn : ST_Recipe;
END_VAR
VAR_OUTPUT
    recipeAdded : BOOL;
    recipeDeleted : BOOL;
    recipeModified : BOOL;
    recipeQueryResult : ST_Recipe;
    error : BOOL;
    status : WORD;
END_VAR
VAR_IN_OUT
    recipe : ARRAY[1..10] OF ST_Recipe;
END_VAR
VAR
    tmp_i : INT;
    tmp_idx : INT;
    tmp_empty : INT;
    tmp_duplicate : BOOL;
    tmp_count : INT;
END_VAR

(* ENGINEERING_CONTRACT
   Pub outputs recipeAdded/Deleted/Modified are one-scan success pulses; no latch.
   error/status are combinational: FALSE/0 on success or idle, TRUE/code on specified failure.
   recipe array persists in IN_OUT slots. Add uses first empty slot; delete clears ID only; modify replaces whole recipe.
   Query/delete/modify search only non-zero recipeID; add duplicate check includes recipeID 0 as empty-slot duplicate.
   Multiple simultaneous request inputs are unspecified; implementation reports error=TRUE, status=16#8000 and performs none.
   Boundary: recipeID 0 is never a queryable/deletable/modifiable identifier.
*)
(* CONTRACT_RULES [] *)

recipeAdded := FALSE;
recipeDeleted := FALSE;
recipeModified := FALSE;
error := FALSE;
status := 0;
recipeQueryResult.recipeID := 0;
recipeQueryResult.ingredientType := 0;
recipeQueryResult.ingredientRatio := 0.0;
recipeQueryResult.productionTemperature := 0.0;

tmp_count := 0;
IF addRecipe THEN
    tmp_count := tmp_count + 1;
END_IF;
IF deleteRecipe THEN
    tmp_count := tmp_count + 1;
END_IF;
IF modifyRecipe THEN
    tmp_count := tmp_count + 1;
END_IF;
IF queryRecipe THEN
    tmp_count := tmp_count + 1;
END_IF;

IF tmp_count > 1 THEN
    error := TRUE;
    status := 16#8000;
    RETURN;
END_IF;

IF addRecipe THEN
    tmp_duplicate := FALSE;
    FOR tmp_i := 1 TO 10 DO
        IF recipe[tmp_i].recipeID = recipeIn.recipeID THEN
            tmp_duplicate := TRUE;
            EXIT;
        END_IF;
    END_FOR;

    IF tmp_duplicate THEN
        error := TRUE;
        status := 16#8002;
    ELSE
        tmp_empty := 0;
        FOR tmp_i := 1 TO 10 DO
            IF recipe[tmp_i].recipeID = 0 THEN
                tmp_empty := tmp_i;
                EXIT;
            END_IF;
        END_FOR;

        IF tmp_empty = 0 THEN
            error := TRUE;
            status := 16#8003;
        ELSE
            recipe[tmp_empty] := recipeIn;
            recipeAdded := TRUE;
        END_IF;
    END_IF;

ELSIF deleteRecipe THEN
    tmp_idx := 0;
    IF recipeIn.recipeID <> 0 THEN
        FOR tmp_i := 1 TO 10 DO
            IF recipe[tmp_i].recipeID = recipeIn.recipeID THEN
                tmp_idx := tmp_i;
                EXIT;
            END_IF;
        END_FOR;
    END_IF;

    IF tmp_idx = 0 THEN
        error := TRUE;
        status := 16#8004;
    ELSE
        recipe[tmp_idx].recipeID := 0;
        recipeDeleted := TRUE;
    END_IF;

ELSIF modifyRecipe THEN
    tmp_idx := 0;
    IF recipeIn.recipeID <> 0 THEN
        FOR tmp_i := 1 TO 10 DO
            IF recipe[tmp_i].recipeID = recipeIn.recipeID THEN
                tmp_idx := tmp_i;
                EXIT;
            END_IF;
        END_FOR;
    END_IF;

    IF tmp_idx = 0 THEN
        error := TRUE;
        status := 16#8005;
    ELSE
        recipe[tmp_idx] := recipeIn;
        recipeModified := TRUE;
    END_IF;

ELSIF queryRecipe THEN
    tmp_idx := 0;
    IF recipeIn.recipeID <> 0 THEN
        FOR tmp_i := 1 TO 10 DO
            IF recipe[tmp_i].recipeID = recipeIn.recipeID THEN
                tmp_idx := tmp_i;
                EXIT;
            END_IF;
        END_FOR;
    END_IF;

    IF tmp_idx = 0 THEN
        error := TRUE;
        status := 16#8001;
    ELSE
        recipeQueryResult := recipe[tmp_idx];
    END_IF;
END_IF;

(* ---- public-hard-03.raw_candidate_02.st ---- *)
TYPE ST_Recipe :
STRUCT
    recipeID : INT;
    ingredientType : INT;
    ingredientRatio : REAL;
    productionTemperature : REAL;
END_STRUCT
END_TYPE;

FUNCTION_BLOCK RecipeManagement
VAR_INPUT
    addRecipe : BOOL;
    deleteRecipe : BOOL;
    modifyRecipe : BOOL;
    queryRecipe : BOOL;
    recipeIn : ST_Recipe;
END_VAR
VAR_OUTPUT
    recipeAdded : BOOL;
    recipeDeleted : BOOL;
    recipeModified : BOOL;
    recipeQueryResult : ST_Recipe;
    error : BOOL;
    status : WORD;
END_VAR
VAR_IN_OUT
    recipe : ARRAY[1..10] OF ST_Recipe;
END_VAR
VAR
    tmp_i : INT;
    tmp_idx : INT;
    tmp_empty : INT;
    tmp_duplicate : BOOL;
    tmp_count : INT;
END_VAR

(* ENGINEERING_CONTRACT
   Pub outputs recipeAdded/Deleted/Modified are one-scan success pulses; no latch.
   error/status are combinational: FALSE/0 on success or idle, TRUE/code on specified failure.
   recipe array persists in IN_OUT slots. Add uses first empty slot; delete clears ID only; modify replaces whole recipe.
   Query/delete/modify search only non-zero recipeID; add duplicate check includes recipeID 0 as empty-slot duplicate.
   Multiple simultaneous request inputs are unspecified; implementation reports error=TRUE, status=16#8000 and performs none.
   Boundary: recipeID 0 is never a queryable/deletable/modifiable identifier.
*)
(* CONTRACT_RULES [] *)

recipeAdded := FALSE;
recipeDeleted := FALSE;
recipeModified := FALSE;
error := FALSE;
status := 0;
recipeQueryResult.recipeID := 0;
recipeQueryResult.ingredientType := 0;
recipeQueryResult.ingredientRatio := 0.0;
recipeQueryResult.productionTemperature := 0.0;

tmp_count := 0;
IF addRecipe THEN
    tmp_count := tmp_count + 1;
END_IF;
IF deleteRecipe THEN
    tmp_count := tmp_count + 1;
END_IF;
IF modifyRecipe THEN
    tmp_count := tmp_count + 1;
END_IF;
IF queryRecipe THEN
    tmp_count := tmp_count + 1;
END_IF;

IF tmp_count > 1 THEN
    error := TRUE;
    status := 16#8000;
    RETURN;
END_IF;

IF addRecipe THEN
    tmp_duplicate := FALSE;
    FOR tmp_i := 1 TO 10 DO
        IF recipe[tmp_i].recipeID = recipeIn.recipeID THEN
            tmp_duplicate := TRUE;
            EXIT;
        END_IF;
    END_FOR;

    IF tmp_duplicate THEN
        error := TRUE;
        status := 16#8002;
    ELSE
        tmp_empty := 0;
        FOR tmp_i := 1 TO 10 DO
            IF recipe[tmp_i].recipeID = 0 THEN
                tmp_empty := tmp_i;
                EXIT;
            END_IF;
        END_FOR;

        IF tmp_empty = 0 THEN
            error := TRUE;
            status := 16#8003;
        ELSE
            recipe[tmp_empty] := recipeIn;
            recipeAdded := TRUE;
        END_IF;
    END_IF;

ELSIF deleteRecipe THEN
    tmp_idx := 0;
    IF recipeIn.recipeID <> 0 THEN
        FOR tmp_i := 1 TO 10 DO
            IF recipe[tmp_i].recipeID = recipeIn.recipeID THEN
                tmp_idx := tmp_i;
                EXIT;
            END_IF;
        END_FOR;
    END_IF;

    IF tmp_idx = 0 THEN
        error := TRUE;
        status := 16#8004;
    ELSE
        recipe[tmp_idx].recipeID := 0;
        recipeDeleted := TRUE;
    END_IF;

ELSIF modifyRecipe THEN
    tmp_idx := 0;
    IF recipeIn.recipeID <> 0 THEN
        FOR tmp_i := 1 TO 10 DO
            IF recipe[tmp_i].recipeID = recipeIn.recipeID THEN
                tmp_idx := tmp_i;
                EXIT;
            END_IF;
        END_FOR;
    END_IF;

    IF tmp_idx = 0 THEN
        error := TRUE;
        status := 16#8005;
    ELSE
        recipe[tmp_idx] := recipeIn;
        recipeModified := TRUE;
    END_IF;

ELSIF queryRecipe THEN
    tmp_idx := 0;
    IF recipeIn.recipeID <> 0 THEN
        FOR tmp_i := 1 TO 10 DO
            IF recipe[tmp_i].recipeID = recipeIn.recipeID THEN
                tmp_idx := tmp_i;
                EXIT;
            END_IF;
        END_FOR;
    END_IF;

    IF tmp_idx = 0 THEN
        error := TRUE;
        status := 16#8001;
    ELSE
        recipeQueryResult := recipe[tmp_idx];
    END_IF;
END_IF;

END_FUNCTION_BLOCK

(* ---- public-hard-03.raw_candidate_03.st ---- *)
TYPE ST_Recipe :
STRUCT
    recipeID : INT;
    ingredientType : INT;
    ingredientRatio : REAL;
    productionTemperature : REAL;
END_STRUCT
END_TYPE;

FUNCTION_BLOCK RecipeManagement
VAR_INPUT
    addRecipe : BOOL;
    deleteRecipe : BOOL;
    modifyRecipe : BOOL;
    queryRecipe : BOOL;
    recipeIn : ST_Recipe;
END_VAR
VAR_OUTPUT
    recipeAdded : BOOL;
    recipeDeleted : BOOL;
    recipeModified : BOOL;
    recipeQueryResult : ST_Recipe;
    error : BOOL;
    status : WORD;
END_VAR
VAR_IN_OUT
    recipe : ARRAY[1..10] OF ST_Recipe;
END_VAR
VAR
    trg_add : R_TRIG;
    trg_delete : R_TRIG;
    trg_modify : R_TRIG;
    trg_query : R_TRIG;
    tmp_i : INT;
    tmp_idx : INT;
    tmp_empty : INT;
    tmp_duplicate : BOOL;
    tmp_count : INT;
END_VAR

(* ENGINEERING_CONTRACT
   Pub outputs recipeAdded/Deleted/Modified are one-scan success pulses; no latch.
   error/status are combinational: FALSE/0 on success or idle, TRUE/code on specified failure.
   recipe array persists in IN_OUT slots. Add uses first empty slot; delete clears ID only; modify replaces whole recipe.
   Query/delete/modify search only non-zero recipeID; add duplicate check includes recipeID 0 as empty-slot duplicate.
   Multiple simultaneous request inputs are unspecified; implementation reports error=TRUE, status=16#8000 and performs none.
   Boundary: recipeID 0 is never a queryable/deletable/modifiable identifier.
*)
(* CONTRACT_RULES [] *)

trg_add(CLK := addRecipe);
trg_delete(CLK := deleteRecipe);
trg_modify(CLK := modifyRecipe);
trg_query(CLK := queryRecipe);

recipeAdded := FALSE;
recipeDeleted := FALSE;
recipeModified := FALSE;
error := FALSE;
status := 0;
recipeQueryResult.recipeID := 0;
recipeQueryResult.ingredientType := 0;
recipeQueryResult.ingredientRatio := 0.0;
recipeQueryResult.productionTemperature := 0.0;

tmp_count := 0;
IF trg_add.Q THEN
    tmp_count := tmp_count + 1;
END_IF;
IF trg_delete.Q THEN
    tmp_count := tmp_count + 1;
END_IF;
IF trg_modify.Q THEN
    tmp_count := tmp_count + 1;
END_IF;
IF trg_query.Q THEN
    tmp_count := tmp_count + 1;
END_IF;

IF tmp_count > 1 THEN
    error := TRUE;
    status := 16#8000;
    RETURN;
END_IF;

IF trg_add.Q THEN
    tmp_duplicate := FALSE;
    FOR tmp_i := 1 TO 10 DO
        IF recipe[tmp_i].recipeID = recipeIn.recipeID THEN
            tmp_duplicate := TRUE;
            EXIT;
        END_IF;
    END_FOR;

    IF tmp_duplicate THEN
        error := TRUE;
        status := 16#8002;
    ELSE
        tmp_empty := 0;
        FOR tmp_i := 1 TO 10 DO
            IF recipe[tmp_i].recipeID = 0 THEN
                tmp_empty := tmp_i;
                EXIT;
            END_IF;
        END_FOR;

        IF tmp_empty = 0 THEN
            error := TRUE;
            status := 16#8003;
        ELSE
            recipe[tmp_empty] := recipeIn;
            recipeAdded := TRUE;
        END_IF;
    END_IF;

ELSIF trg_delete.Q THEN
    tmp_idx := 0;
    IF recipeIn.recipeID <> 0 THEN
        FOR tmp_i := 1 TO 10 DO
            IF recipe[tmp_i].recipeID = recipeIn.recipeID THEN
                tmp_idx := tmp_i;
                EXIT;
            END_IF;
        END_FOR;
    END_IF;

    IF tmp_idx = 0 THEN
        error := TRUE;
        status := 16#8004;
    ELSE
        recipe[tmp_idx].recipeID := 0;
        recipeDeleted := TRUE;
    END_IF;

ELSIF trg_modify.Q THEN
    tmp_idx := 0;
    IF recipeIn.recipeID <> 0 THEN
        FOR tmp_i := 1 TO 10 DO
            IF recipe[tmp_i].recipeID = recipeIn.recipeID THEN
                tmp_idx := tmp_i;
                EXIT;
            END_IF;
        END_FOR;
    END_IF;

    IF tmp_idx = 0 THEN
        error := TRUE;
        status := 16#8005;
    ELSE
        recipe[tmp_idx] := recipeIn;
        recipeModified := TRUE;
    END_IF;

ELSIF trg_query.Q THEN
    tmp_idx := 0;
    IF recipeIn.recipeID <> 0 THEN
        FOR tmp_i := 1 TO 10 DO
            IF recipe[tmp_i].recipeID = recipeIn.recipeID THEN
                tmp_idx := tmp_i;
                EXIT;
            END_IF;
        END_FOR;
    END_IF;

    IF tmp_idx = 0 THEN
        error := TRUE;
        status := 16#8001;
    ELSE
        recipeQueryResult := recipe[tmp_idx];
    END_IF;
END_IF;

END_FUNCTION_BLOCK

(* ---- public-hard-03.raw_candidate_04.st ---- *)
TYPE ST_Recipe :
STRUCT
    recipeID : INT;
    ingredientType : INT;
    ingredientRatio : REAL;
    productionTemperature : REAL;
END_STRUCT
END_TYPE;

FUNCTION_BLOCK RecipeManagement
VAR_INPUT
    addRecipe : BOOL;
    deleteRecipe : BOOL;
    modifyRecipe : BOOL;
    queryRecipe : BOOL;
    recipeIn : ST_Recipe;
END_VAR
VAR_OUTPUT
    recipeAdded : BOOL;
    recipeDeleted : BOOL;
    recipeModified : BOOL;
    recipeQueryResult : ST_Recipe;
    error : BOOL;
    status : WORD;
END_VAR
VAR_IN_OUT
    recipe : ARRAY[1..10] OF ST_Recipe;
END_VAR
VAR
    trg_add : R_TRIG;
    trg_delete : R_TRIG;
    trg_modify : R_TRIG;
    trg_query : R_TRIG;
    tmp_i : INT;
    tmp_idx : INT;
    tmp_empty : INT;
    tmp_duplicate : BOOL;
    tmp_count : INT;
END_VAR

(* ENGINEERING_CONTRACT
   Pub outputs recipeAdded/Deleted/Modified are one-scan success pulses; no latch.
   error/status are combinational: FALSE/0 on success or idle, TRUE/code on specified failure.
   recipe array persists in IN_OUT slots. Add uses first empty slot; delete clears ID only; modify replaces whole recipe.
   Query/delete/modify search only non-zero recipeID; add duplicate check includes recipeID 0 as empty-slot duplicate.
   Multiple simultaneous request inputs are unspecified; implementation reports error=TRUE, status=16#8000 and performs none.
   Boundary: recipeID 0 is never a queryable/deletable/modifiable identifier.
   recipeQueryResult is retained after a successful query until the next successful query. It is not cleared on idle or on an unsuccessful query.
*)
(* CONTRACT_RULES [] *)

trg_add(CLK := addRecipe);
trg_delete(CLK := deleteRecipe);
trg_modify(CLK := modifyRecipe);
trg_query(CLK := queryRecipe);

recipeAdded := FALSE;
recipeDeleted := FALSE;
recipeModified := FALSE;
error := FALSE;
status := 0;

tmp_count := 0;
IF trg_add.Q THEN
    tmp_count := tmp_count + 1;
END_IF;
IF trg_delete.Q THEN
    tmp_count := tmp_count + 1;
END_IF;
IF trg_modify.Q THEN
    tmp_count := tmp_count + 1;
END_IF;
IF trg_query.Q THEN
    tmp_count := tmp_count + 1;
END_IF;

IF tmp_count > 1 THEN
    error := TRUE;
    status := 16#8000;
    RETURN;
END_IF;

IF trg_add.Q THEN
    tmp_duplicate := FALSE;
    FOR tmp_i := 1 TO 10 DO
        IF recipe[tmp_i].recipeID = recipeIn.recipeID THEN
            tmp_duplicate := TRUE;
            EXIT;
        END_IF;
    END_FOR;

    IF tmp_duplicate THEN
        error := TRUE;
        status := 16#8002;
    ELSE
        tmp_empty := 0;
        FOR tmp_i := 1 TO 10 DO
            IF recipe[tmp_i].recipeID = 0 THEN
                tmp_empty := tmp_i;
                EXIT;
            END_IF;
        END_FOR;

        IF tmp_empty = 0 THEN
            error := TRUE;
            status := 16#8003;
        ELSE
            recipe[tmp_empty] := recipeIn;
            recipeAdded := TRUE;
        END_IF;
    END_IF;

ELSIF trg_delete.Q THEN
    tmp_idx := 0;
    IF recipeIn.recipeID <> 0 THEN
        FOR tmp_i := 1 TO 10 DO
            IF recipe[tmp_i].recipeID = recipeIn.recipeID THEN
                tmp_idx := tmp_i;
                EXIT;
            END_IF;
        END_FOR;
    END_IF;

    IF tmp_idx = 0 THEN
        error := TRUE;
        status := 16#8004;
    ELSE
        recipe[tmp_idx].recipeID := 0;
        recipeDeleted := TRUE;
    END_IF;

ELSIF trg_modify.Q THEN
    tmp_idx := 0;
    IF recipeIn.recipeID <> 0 THEN
        FOR tmp_i := 1 TO 10 DO
            IF recipe[tmp_i].recipeID = recipeIn.recipeID THEN
                tmp_idx := tmp_i;
                EXIT;
            END_IF;
        END_FOR;
    END_IF;

    IF tmp_idx = 0 THEN
        error := TRUE;
        status := 16#8005;
    ELSE
        recipe[tmp_idx] := recipeIn;
        recipeModified := TRUE;
    END_IF;

ELSIF trg_query.Q THEN
    tmp_idx := 0;
    IF recipeIn.recipeID <> 0 THEN
        FOR tmp_i := 1 TO 10 DO
            IF recipe[tmp_i].recipeID = recipeIn.recipeID THEN
                tmp_idx := tmp_i;
                EXIT;
            END_IF;
        END_FOR;
    END_IF;

    IF tmp_idx = 0 THEN
        error := TRUE;
        status := 16#8001;
    ELSE
        recipeQueryResult := recipe[tmp_idx];
    END_IF;
END_IF;

END_FUNCTION_BLOCK

(* ---- public-hard-04.candidate_01.st ---- *)
(* ENGINEERING_CONTRACT
   elementCount DINT: retained process value; 0 after reset, +1 successful enqueue, -1 successful dequeue, held otherwise; range 0..capacity.
   status WORD: overwritten every invocation; 0 idle/reset/success, 16#8002 rejected full enqueue, 16#8001 rejected empty dequeue; reset priority sets 0.
   queue state: first invocation empty; reset priority clears head/tail/count; enqueue writes at tail, dequeue reads head; indices 0..capacity-1.
   edge triggers: R_TRIG consumed every scan; reset priority ignores edge requests; simultaneous enqueue+dequeue unspecified -> no-op.
   units/boundaries: capacity positive DINT derived once from buffer size / item element size; element copied byte-wise from item address.
*)
(* CONTRACT_RULES [] *)
FUNCTION_BLOCK FIFO
VAR_INPUT
    enqueue : BOOL;
    dequeue : BOOL;
    reset : BOOL;
END_VAR
VAR_OUTPUT
    elementCount : DINT;
    status : WORD;
END_VAR
VAR_IN_OUT
    item : VARIANT;
    buffer : VARIANT;
END_VAR
VAR
    local_rEnq : R_TRIG;
    local_rDeq : R_TRIG;
    local_enqEdge : BOOL;
    local_deqEdge : BOOL;

    local_associated : BOOL := FALSE;
    local_pBufferBase : POINTER TO BYTE;
    local_pItemBase : POINTER TO BYTE;
    local_elemSize : DINT := 1;
    local_capacity : DINT := 1;

    local_count : DINT := 0;
    local_head : DINT := 0;
    local_tail : DINT := 0;

    local_bufInfo : __SYSTEM.VAR_INFO;
    local_itemInfo : __SYSTEM.VAR_INFO;

    local_pSrc : POINTER TO BYTE;
    local_pDst : POINTER TO BYTE;
    local_i : DINT;
END_VAR

(* Consume rising edges every scan so reset cannot create ghost operations later. *)
local_rEnq(CLK := enqueue);
local_enqEdge := local_rEnq.Q;
local_rDeq(CLK := dequeue);
local_deqEdge := local_rDeq.Q;

status := 16#0000;

(* One-time association of buffer and element storage, using the first invocation. *)
IF NOT local_associated THEN
    local_bufInfo := __VARINFO(buffer);
    local_itemInfo := __VARINFO(item);

    local_elemSize := local_itemInfo.diSize;
    IF local_elemSize <= 0 THEN
        local_elemSize := 1;
    END_IF;

    local_capacity := local_bufInfo.diSize / local_elemSize;
    IF local_capacity < 1 THEN
        local_capacity := 1;
    END_IF;

    local_pBufferBase := local_bufInfo.pvAddress;
    local_pItemBase := local_itemInfo.pvAddress;
    local_associated := TRUE;
END_IF;

IF reset THEN
    (* Reset has priority over all operations; stored values remain untouched. *)
    local_count := 0;
    local_head := 0;
    local_tail := 0;
    status := 16#0000;
ELSE
    IF local_enqEdge AND NOT local_deqEdge THEN
        IF local_count < local_capacity THEN
            (* Copy current item value into tail slot. *)
            local_pSrc := local_pItemBase;
            local_pDst := local_pBufferBase + (local_tail * local_elemSize);

            FOR local_i := 0 TO local_elemSize - 1 DO
                local_pDst^ := local_pSrc^;
                local_pSrc := local_pSrc + 1;
                local_pDst := local_pDst + 1;
            END_FOR;

            local_tail := (local_tail + 1) MOD local_capacity;
            local_count := local_count + 1;
            status := 16#0000;
        ELSE
            status := 16#8002; (* enqueue rejected: full *)
        END_IF;
    ELSIF local_deqEdge AND NOT local_enqEdge THEN
        IF local_count > 0 THEN
            (* Copy head element back to item. *)
            local_pSrc := local_pBufferBase + (local_head * local_elemSize);
            local_pDst := local_pItemBase;

            FOR local_i := 0 TO local_elemSize - 1 DO
                local_pDst^ := local_pSrc^;
                local_pSrc := local_pSrc + 1;
                local_pDst := local_pDst + 1;
            END_FOR;

            local_head := (local_head + 1) MOD local_capacity;
            local_count := local_count - 1;
            status := 16#0000;
        ELSE
            status := 16#8001; (* dequeue rejected: empty *)
        END_IF;
    END_IF;
END_IF;

elementCount := local_count;

(* ---- public-hard-04.candidate_02.st ---- *)
(* ENGINEERING_CONTRACT
   elementCount DINT: retained process value; 0 after reset, +1 successful enqueue, -1 successful dequeue, held otherwise; range 0..capacity.
   status WORD: overwritten every invocation; 0 idle/reset/success, 16#8002 rejected full enqueue, 16#8001 rejected empty dequeue; reset priority sets 0.
   queue state: first invocation empty; reset priority clears head/tail/count; enqueue writes at tail, dequeue reads head; indices 0..capacity-1.
   edge triggers: R_TRIG consumed every scan; reset priority ignores edge requests; simultaneous enqueue+dequeue unspecified -> no-op.
   units/boundaries: capacity positive DINT derived once from buffer size / item element size; element copied byte-wise from item address.
*)
(* CONTRACT_RULES [] *)
FUNCTION_BLOCK FIFO
VAR_INPUT
    enqueue : BOOL;
    dequeue : BOOL;
    reset : BOOL;
END_VAR
VAR_OUTPUT
    elementCount : DINT;
    status : WORD;
END_VAR
VAR_IN_OUT
    item : VARIANT;
    buffer : VARIANT;
END_VAR
VAR
    local_rEnq : R_TRIG;
    local_rDeq : R_TRIG;
    local_enqEdge : BOOL;
    local_deqEdge : BOOL;

    local_associated : BOOL := FALSE;
    local_pBufferBase : POINTER TO BYTE;
    local_pItemBase : POINTER TO BYTE;
    local_elemSize : DINT := 1;
    local_capacity : DINT := 1;

    local_count : DINT := 0;
    local_head : DINT := 0;
    local_tail : DINT := 0;

    local_bufInfo : __SYSTEM.VAR_INFO;
    local_itemInfo : __SYSTEM.VAR_INFO;

    local_pSrc : POINTER TO BYTE;
    local_pDst : POINTER TO BYTE;
    local_offset : DINT;
    local_copiedBytes : UDINT;
END_VAR

(* Consume rising edges every scan so reset cannot create ghost operations later. *)
local_rEnq(CLK := enqueue);
local_enqEdge := local_rEnq.Q;
local_rDeq(CLK := dequeue);
local_deqEdge := local_rDeq.Q;

status := 16#0000;

(* One-time association of buffer and item storage, using the first invocation. *)
IF NOT local_associated THEN
    local_bufInfo := __VARINFO(buffer);
    local_itemInfo := __VARINFO(item);

    local_elemSize := local_itemInfo.diSize;
    IF local_elemSize <= 0 THEN
        local_elemSize := 1;
    END_IF;

    local_capacity := local_bufInfo.diSize / local_elemSize;
    IF local_capacity < 1 THEN
        local_capacity := 1;
    END_IF;

    local_pBufferBase := local_bufInfo.pvAddress;
    local_pItemBase := local_itemInfo.pvAddress;
    local_associated := TRUE;
END_IF;

IF reset THEN
    (* Reset has priority over all operations; stored values remain untouched. *)
    local_count := 0;
    local_head := 0;
    local_tail := 0;
    status := 16#0000;
ELSE
    IF local_enqEdge AND NOT local_deqEdge THEN
        IF local_count < local_capacity THEN
            (* Copy current item value into tail slot. *)
            local_pSrc := local_pItemBase;
            local_pDst := local_pBufferBase;
            local_offset := local_tail * local_elemSize;
            local_pDst := local_pDst + local_offset;
            local_copiedBytes := SysMemCpy(
                pbyDest := local_pDst,
                pbySource := local_pSrc,
                dwCount := TO_DWORD(local_elemSize)
            );

            local_tail := (local_tail + 1) MOD local_capacity;
            local_count := local_count + 1;
            status := 16#0000;
        ELSE
            status := 16#8002; (* enqueue rejected: full *)
        END_IF;
    ELSIF local_deqEdge AND NOT local_enqEdge THEN
        IF local_count > 0 THEN
            (* Copy head element back to item. *)
            local_pSrc := local_pBufferBase;
            local_offset := local_head * local_elemSize;
            local_pSrc := local_pSrc + local_offset;
            local_pDst := local_pItemBase;
            local_copiedBytes := SysMemCpy(
                pbyDest := local_pDst,
                pbySource := local_pSrc,
                dwCount := TO_DWORD(local_elemSize)
            );

            local_head := (local_head + 1) MOD local_capacity;
            local_count := local_count - 1;
            status := 16#0000;
        ELSE
            status := 16#8001; (* dequeue rejected: empty *)
        END_IF;
    END_IF;
END_IF;

elementCount := local_count;

(* ---- public-hard-04.candidate_03.st ---- *)
(* ENGINEERING_CONTRACT
   elementCount DINT: retained process value; 0 after reset, +1 successful enqueue, -1 successful dequeue, held otherwise; range 0..capacity.
   status WORD: overwritten every invocation; 0 idle/reset/success, 16#8002 rejected full enqueue, 16#8001 rejected empty dequeue; reset priority sets 0.
   queue state: first invocation empty; reset priority clears head/tail/count; enqueue writes at tail, dequeue reads head; indices 0..capacity-1.
   edge triggers: R_TRIG consumed every scan; reset priority ignores edge requests; simultaneous enqueue+dequeue unspecified -> no-op.
   units/boundaries: capacity positive DINT derived once from buffer size / item element size; element copied byte-wise from item address.
*)
(* CONTRACT_RULES [] *)
FUNCTION_BLOCK FIFO
VAR_INPUT
    enqueue : BOOL;
    dequeue : BOOL;
    reset : BOOL;
END_VAR
VAR_OUTPUT
    elementCount : DINT;
    status : WORD;
END_VAR
VAR_IN_OUT
    item : VARIANT;
    buffer : VARIANT;
END_VAR
VAR
    local_rEnq : R_TRIG;
    local_rDeq : R_TRIG;
    local_enqEdge : BOOL;
    local_deqEdge : BOOL;

    local_associated : BOOL := FALSE;
    local_pBufferBase : POINTER TO BYTE;
    local_pItemBase : POINTER TO BYTE;
    local_elemSize : DINT := 1;
    local_capacity : DINT := 1;

    local_count : DINT := 0;
    local_head : DINT := 0;
    local_tail : DINT := 0;

    local_bufInfo : __SYSTEM.VAR_INFO;
    local_itemInfo : __SYSTEM.VAR_INFO;

    local_pSrc : POINTER TO BYTE;
    local_pDst : POINTER TO BYTE;
    local_offset : DINT;
    local_copiedBytes : UDINT;
END_VAR

(* Consume rising edges every scan so reset cannot create ghost operations later. *)
local_rEnq(CLK := enqueue);
local_enqEdge := local_rEnq.Q;
local_rDeq(CLK := dequeue);
local_deqEdge := local_rDeq.Q;

status := 16#0000;

(* One-time association of buffer and item storage, using the first invocation. *)
IF NOT local_associated THEN
    local_bufInfo := __VARINFO(buffer);
    local_itemInfo := __VARINFO(item);

    local_elemSize := local_itemInfo.diSize;
    IF local_elemSize <= 0 THEN
        local_elemSize := 1;
    END_IF;

    local_capacity := local_bufInfo.diSize / local_elemSize;
    IF local_capacity < 1 THEN
        local_capacity := 1;
    END_IF;

    local_pBufferBase := local_bufInfo.pvAddress;
    local_pItemBase := local_itemInfo.pvAddress;
    local_associated := TRUE;
END_IF;

IF reset THEN
    (* Reset has priority over all operations; stored values remain untouched. *)
    local_count := 0;
    local_head := 0;
    local_tail := 0;
    status := 16#0000;
ELSE
    IF local_enqEdge AND NOT local_deqEdge THEN
        IF local_count < local_capacity THEN
            (* Copy current item value into tail slot. *)
            local_pSrc := local_pItemBase;
            local_pDst := local_pBufferBase;
            local_offset := local_tail * local_elemSize;
            local_pDst := local_pDst + local_offset;
            local_copiedBytes := SysMemCpy(
                pbyDest := local_pDst,
                pbySource := local_pSrc,
                dwCount := TO_DWORD(local_elemSize)
            );

            local_tail := (local_tail + 1) MOD local_capacity;
            local_count := local_count + 1;
            status := 16#0000;
        ELSE
            status := 16#8002; (* enqueue rejected: full *)
        END_IF;
    ELSIF local_deqEdge AND NOT local_enqEdge THEN
        IF local_count > 0 THEN
            (* Copy head element back to item. *)
            local_pSrc := local_pBufferBase;
            local_offset := local_head * local_elemSize;
            local_pSrc := local_pSrc + local_offset;
            local_pDst := local_pItemBase;
            local_copiedBytes := SysMemCpy(
                pbyDest := local_pDst,
                pbySource := local_pSrc,
                dwCount := TO_DWORD(local_elemSize)
            );

            local_head := (local_head + 1) MOD local_capacity;
            local_count := local_count - 1;
            status := 16#0000;
        ELSE
            status := 16#8001; (* dequeue rejected: empty *)
        END_IF;
    END_IF;
END_IF;

elementCount := local_count;
END_FUNCTION_BLOCK

(* ---- public-hard-04.candidate_04.st ---- *)
(* ENGINEERING_CONTRACT
   elementCount DINT: retained process value; 0 after reset, +1 successful enqueue, -1 successful dequeue, held otherwise; range 0..capacity.
   status WORD: overwritten every invocation; 0 idle/reset/success, 16#8002 rejected full enqueue, 16#8001 rejected empty dequeue; reset priority sets 0.
   queue state: first invocation empty; reset priority clears head/tail/count; enqueue writes at tail, dequeue reads head; indices 0..capacity-1.
   edge triggers: R_TRIG consumed every scan; reset priority ignores edge requests; simultaneous enqueue+dequeue unspecified -> no-op.
   units/boundaries: capacity positive DINT derived once from buffer size / item element size; element copied byte-wise from item address.
*)
(* CONTRACT_RULES [] *)
FUNCTION_BLOCK FIFO
VAR_INPUT
    enqueue : BOOL;
    dequeue : BOOL;
    reset : BOOL;
END_VAR
VAR_OUTPUT
    elementCount : DINT;
    status : WORD;
END_VAR
VAR_IN_OUT
    item : VARIANT;
    buffer : VARIANT;
END_VAR
VAR
    local_rEnq : R_TRIG;
    local_rDeq : R_TRIG;
    local_enqEdge : BOOL;
    local_deqEdge : BOOL;

    local_associated : BOOL := FALSE;
    local_pBufferBase : POINTER TO BYTE;
    local_pItemBase : POINTER TO BYTE;
    local_elemSize : DINT := 1;
    local_capacity : DINT := 1;

    local_count : DINT := 0;
    local_head : DINT := 0;
    local_tail : DINT := 0;

    local_bufInfo : __SYSTEM.VAR_INFO;
    local_itemInfo : __SYSTEM.VAR_INFO;

    local_pSrc : POINTER TO BYTE;
    local_pDst : POINTER TO BYTE;
    local_offset : DINT;
    local_copiedBytes : UDINT;
END_VAR

(* Consume rising edges every scan so reset cannot create ghost operations later. *)
local_rEnq(CLK := enqueue);
local_enqEdge := local_rEnq.Q;
local_rDeq(CLK := dequeue);
local_deqEdge := local_rDeq.Q;

status := 16#0000;

(* One-time association of buffer and item storage, using the first invocation. *)
IF NOT local_associated THEN
    local_bufInfo := __VARINFO(buffer);
    local_itemInfo := __VARINFO(item);

    local_elemSize := local_itemInfo.diSize;
    IF local_elemSize <= 0 THEN
        local_elemSize := 1;
    END_IF;

    local_capacity := local_bufInfo.diSize / local_elemSize;
    IF local_capacity < 1 THEN
        local_capacity := 1;
    END_IF;

    local_pBufferBase := local_bufInfo.pvAddress;
    local_pItemBase := local_itemInfo.pvAddress;
    local_associated := TRUE;
END_IF;

IF reset THEN
    (* Reset has priority over all operations; stored values remain untouched. *)
    local_count := 0;
    local_head := 0;
    local_tail := 0;
    status := 16#0000;
ELSE
    IF local_enqEdge AND NOT local_deqEdge THEN
        IF local_count < local_capacity THEN
            (* Copy current item value into tail slot. *)
            local_pSrc := local_pItemBase;
            local_pDst := local_pBufferBase;
            local_offset := local_tail * local_elemSize;
            local_pDst := local_pDst + local_offset;
            local_copiedBytes := SysMemCpy(
                pbyDest := local_pDst,
                pbySource := local_pSrc,
                dwCount := TO_DWORD(local_elemSize)
            );

            local_tail := (local_tail + 1) MOD local_capacity;
            local_count := local_count + 1;
            status := 16#0000;
        ELSE
            status := 16#8002; (* enqueue rejected: full *)
        END_IF;
    ELSIF local_deqEdge AND NOT local_enqEdge THEN
        IF local_count > 0 THEN
            (* Copy head element back to item. *)
            local_pSrc := local_pBufferBase;
            local_offset := local_head * local_elemSize;
            local_pSrc := local_pSrc + local_offset;
            local_pDst := local_pItemBase;
            local_copiedBytes := SysMemCpy(
                pbyDest := local_pDst,
                pbySource := local_pSrc,
                dwCount := TO_DWORD(local_elemSize)
            );

            local_head := (local_head + 1) MOD local_capacity;
            local_count := local_count - 1;
            status := 16#0000;
        ELSE
            status := 16#8001; (* dequeue rejected: empty *)
        END_IF;
    END_IF;
END_IF;

elementCount := local_count;
END_FUNCTION_BLOCK

(* ---- public-hard-04.raw_candidate_01.st ---- *)
(* ENGINEERING_CONTRACT
   elementCount DINT: retained process value; 0 after reset, +1 successful enqueue, -1 successful dequeue, held otherwise; range 0..capacity.
   status WORD: overwritten every invocation; 0 idle/reset/success, 16#8002 rejected full enqueue, 16#8001 rejected empty dequeue; reset priority sets 0.
   queue state: first invocation empty; reset priority clears head/tail/count; enqueue writes at tail, dequeue reads head; indices 0..capacity-1.
   edge triggers: R_TRIG consumed every scan; reset priority ignores edge requests; simultaneous enqueue+dequeue unspecified -> no-op.
   units/boundaries: capacity positive DINT derived once from buffer size / item element size; element copied byte-wise from item address.
*)
(* CONTRACT_RULES [] *)
FUNCTION_BLOCK FIFO
VAR_INPUT
    enqueue : BOOL;
    dequeue : BOOL;
    reset : BOOL;
END_VAR
VAR_OUTPUT
    elementCount : DINT;
    status : WORD;
END_VAR
VAR_IN_OUT
    item : VARIANT;
    buffer : VARIANT;
END_VAR
VAR
    local_rEnq : R_TRIG;
    local_rDeq : R_TRIG;
    local_enqEdge : BOOL;
    local_deqEdge : BOOL;

    local_associated : BOOL := FALSE;
    local_pBufferBase : POINTER TO BYTE;
    local_pItemBase : POINTER TO BYTE;
    local_elemSize : DINT := 1;
    local_capacity : DINT := 1;

    local_count : DINT := 0;
    local_head : DINT := 0;
    local_tail : DINT := 0;

    local_bufInfo : __SYSTEM.VAR_INFO;
    local_itemInfo : __SYSTEM.VAR_INFO;

    local_pSrc : POINTER TO BYTE;
    local_pDst : POINTER TO BYTE;
    local_i : DINT;
END_VAR

(* Consume rising edges every scan so reset cannot create ghost operations later. *)
local_rEnq(CLK := enqueue);
local_enqEdge := local_rEnq.Q;
local_rDeq(CLK := dequeue);
local_deqEdge := local_rDeq.Q;

status := 16#0000;

(* One-time association of buffer and element storage, using the first invocation. *)
IF NOT local_associated THEN
    local_bufInfo := __VARINFO(buffer);
    local_itemInfo := __VARINFO(item);

    local_elemSize := local_itemInfo.diSize;
    IF local_elemSize <= 0 THEN
        local_elemSize := 1;
    END_IF;

    local_capacity := local_bufInfo.diSize / local_elemSize;
    IF local_capacity < 1 THEN
        local_capacity := 1;
    END_IF;

    local_pBufferBase := local_bufInfo.pvAddress;
    local_pItemBase := local_itemInfo.pvAddress;
    local_associated := TRUE;
END_IF;

IF reset THEN
    (* Reset has priority over all operations; stored values remain untouched. *)
    local_count := 0;
    local_head := 0;
    local_tail := 0;
    status := 16#0000;
ELSE
    IF local_enqEdge AND NOT local_deqEdge THEN
        IF local_count < local_capacity THEN
            (* Copy current item value into tail slot. *)
            local_pSrc := local_pItemBase;
            local_pDst := local_pBufferBase + (local_tail * local_elemSize);

            FOR local_i := 0 TO local_elemSize - 1 DO
                local_pDst^ := local_pSrc^;
                local_pSrc := local_pSrc + 1;
                local_pDst := local_pDst + 1;
            END_FOR;

            local_tail := (local_tail + 1) MOD local_capacity;
            local_count := local_count + 1;
            status := 16#0000;
        ELSE
            status := 16#8002; (* enqueue rejected: full *)
        END_IF;
    ELSIF local_deqEdge AND NOT local_enqEdge THEN
        IF local_count > 0 THEN
            (* Copy head element back to item. *)
            local_pSrc := local_pBufferBase + (local_head * local_elemSize);
            local_pDst := local_pItemBase;

            FOR local_i := 0 TO local_elemSize - 1 DO
                local_pDst^ := local_pSrc^;
                local_pSrc := local_pSrc + 1;
                local_pDst := local_pDst + 1;
            END_FOR;

            local_head := (local_head + 1) MOD local_capacity;
            local_count := local_count - 1;
            status := 16#0000;
        ELSE
            status := 16#8001; (* dequeue rejected: empty *)
        END_IF;
    END_IF;
END_IF;

elementCount := local_count;

(* ---- public-hard-04.raw_candidate_02.st ---- *)
(* ENGINEERING_CONTRACT
   elementCount DINT: retained process value; 0 after reset, +1 successful enqueue, -1 successful dequeue, held otherwise; range 0..capacity.
   status WORD: overwritten every invocation; 0 idle/reset/success, 16#8002 rejected full enqueue, 16#8001 rejected empty dequeue; reset priority sets 0.
   queue state: first invocation empty; reset priority clears head/tail/count; enqueue writes at tail, dequeue reads head; indices 0..capacity-1.
   edge triggers: R_TRIG consumed every scan; reset priority ignores edge requests; simultaneous enqueue+dequeue unspecified -> no-op.
   units/boundaries: capacity positive DINT derived once from buffer size / item element size; element copied byte-wise from item address.
*)
(* CONTRACT_RULES [] *)
FUNCTION_BLOCK FIFO
VAR_INPUT
    enqueue : BOOL;
    dequeue : BOOL;
    reset : BOOL;
END_VAR
VAR_OUTPUT
    elementCount : DINT;
    status : WORD;
END_VAR
VAR_IN_OUT
    item : VARIANT;
    buffer : VARIANT;
END_VAR
VAR
    local_rEnq : R_TRIG;
    local_rDeq : R_TRIG;
    local_enqEdge : BOOL;
    local_deqEdge : BOOL;

    local_associated : BOOL := FALSE;
    local_pBufferBase : POINTER TO BYTE;
    local_pItemBase : POINTER TO BYTE;
    local_elemSize : DINT := 1;
    local_capacity : DINT := 1;

    local_count : DINT := 0;
    local_head : DINT := 0;
    local_tail : DINT := 0;

    local_bufInfo : __SYSTEM.VAR_INFO;
    local_itemInfo : __SYSTEM.VAR_INFO;

    local_pSrc : POINTER TO BYTE;
    local_pDst : POINTER TO BYTE;
    local_offset : DINT;
    local_copiedBytes : UDINT;
END_VAR

(* Consume rising edges every scan so reset cannot create ghost operations later. *)
local_rEnq(CLK := enqueue);
local_enqEdge := local_rEnq.Q;
local_rDeq(CLK := dequeue);
local_deqEdge := local_rDeq.Q;

status := 16#0000;

(* One-time association of buffer and item storage, using the first invocation. *)
IF NOT local_associated THEN
    local_bufInfo := __VARINFO(buffer);
    local_itemInfo := __VARINFO(item);

    local_elemSize := local_itemInfo.diSize;
    IF local_elemSize <= 0 THEN
        local_elemSize := 1;
    END_IF;

    local_capacity := local_bufInfo.diSize / local_elemSize;
    IF local_capacity < 1 THEN
        local_capacity := 1;
    END_IF;

    local_pBufferBase := local_bufInfo.pvAddress;
    local_pItemBase := local_itemInfo.pvAddress;
    local_associated := TRUE;
END_IF;

IF reset THEN
    (* Reset has priority over all operations; stored values remain untouched. *)
    local_count := 0;
    local_head := 0;
    local_tail := 0;
    status := 16#0000;
ELSE
    IF local_enqEdge AND NOT local_deqEdge THEN
        IF local_count < local_capacity THEN
            (* Copy current item value into tail slot. *)
            local_pSrc := local_pItemBase;
            local_pDst := local_pBufferBase;
            local_offset := local_tail * local_elemSize;
            local_pDst := local_pDst + local_offset;
            local_copiedBytes := SysMemCpy(
                pbyDest := local_pDst,
                pbySource := local_pSrc,
                dwCount := TO_DWORD(local_elemSize)
            );

            local_tail := (local_tail + 1) MOD local_capacity;
            local_count := local_count + 1;
            status := 16#0000;
        ELSE
            status := 16#8002; (* enqueue rejected: full *)
        END_IF;
    ELSIF local_deqEdge AND NOT local_enqEdge THEN
        IF local_count > 0 THEN
            (* Copy head element back to item. *)
            local_pSrc := local_pBufferBase;
            local_offset := local_head * local_elemSize;
            local_pSrc := local_pSrc + local_offset;
            local_pDst := local_pItemBase;
            local_copiedBytes := SysMemCpy(
                pbyDest := local_pDst,
                pbySource := local_pSrc,
                dwCount := TO_DWORD(local_elemSize)
            );

            local_head := (local_head + 1) MOD local_capacity;
            local_count := local_count - 1;
            status := 16#0000;
        ELSE
            status := 16#8001; (* dequeue rejected: empty *)
        END_IF;
    END_IF;
END_IF;

elementCount := local_count;

(* ---- public-hard-04.raw_candidate_03.st ---- *)
(* ENGINEERING_CONTRACT
   elementCount DINT: retained process value; 0 after reset, +1 successful enqueue, -1 successful dequeue, held otherwise; range 0..capacity.
   status WORD: overwritten every invocation; 0 idle/reset/success, 16#8002 rejected full enqueue, 16#8001 rejected empty dequeue; reset priority sets 0.
   queue state: first invocation empty; reset priority clears head/tail/count; enqueue writes at tail, dequeue reads head; indices 0..capacity-1.
   edge triggers: R_TRIG consumed every scan; reset priority ignores edge requests; simultaneous enqueue+dequeue unspecified -> no-op.
   units/boundaries: capacity positive DINT derived once from buffer size / item element size; element copied byte-wise from item address.
*)
(* CONTRACT_RULES [] *)
FUNCTION_BLOCK FIFO
VAR_INPUT
    enqueue : BOOL;
    dequeue : BOOL;
    reset : BOOL;
END_VAR
VAR_OUTPUT
    elementCount : DINT;
    status : WORD;
END_VAR
VAR_IN_OUT
    item : VARIANT;
    buffer : VARIANT;
END_VAR
VAR
    local_rEnq : R_TRIG;
    local_rDeq : R_TRIG;
    local_enqEdge : BOOL;
    local_deqEdge : BOOL;

    local_associated : BOOL := FALSE;
    local_pBufferBase : POINTER TO BYTE;
    local_pItemBase : POINTER TO BYTE;
    local_elemSize : DINT := 1;
    local_capacity : DINT := 1;

    local_count : DINT := 0;
    local_head : DINT := 0;
    local_tail : DINT := 0;

    local_bufInfo : __SYSTEM.VAR_INFO;
    local_itemInfo : __SYSTEM.VAR_INFO;

    local_pSrc : POINTER TO BYTE;
    local_pDst : POINTER TO BYTE;
    local_offset : DINT;
    local_copiedBytes : UDINT;
END_VAR

(* Consume rising edges every scan so reset cannot create ghost operations later. *)
local_rEnq(CLK := enqueue);
local_enqEdge := local_rEnq.Q;
local_rDeq(CLK := dequeue);
local_deqEdge := local_rDeq.Q;

status := 16#0000;

(* One-time association of buffer and item storage, using the first invocation. *)
IF NOT local_associated THEN
    local_bufInfo := __VARINFO(buffer);
    local_itemInfo := __VARINFO(item);

    local_elemSize := local_itemInfo.diSize;
    IF local_elemSize <= 0 THEN
        local_elemSize := 1;
    END_IF;

    local_capacity := local_bufInfo.diSize / local_elemSize;
    IF local_capacity < 1 THEN
        local_capacity := 1;
    END_IF;

    local_pBufferBase := local_bufInfo.pvAddress;
    local_pItemBase := local_itemInfo.pvAddress;
    local_associated := TRUE;
END_IF;

IF reset THEN
    (* Reset has priority over all operations; stored values remain untouched. *)
    local_count := 0;
    local_head := 0;
    local_tail := 0;
    status := 16#0000;
ELSE
    IF local_enqEdge AND NOT local_deqEdge THEN
        IF local_count < local_capacity THEN
            (* Copy current item value into tail slot. *)
            local_pSrc := local_pItemBase;
            local_pDst := local_pBufferBase;
            local_offset := local_tail * local_elemSize;
            local_pDst := local_pDst + local_offset;
            local_copiedBytes := SysMemCpy(
                pbyDest := local_pDst,
                pbySource := local_pSrc,
                dwCount := TO_DWORD(local_elemSize)
            );

            local_tail := (local_tail + 1) MOD local_capacity;
            local_count := local_count + 1;
            status := 16#0000;
        ELSE
            status := 16#8002; (* enqueue rejected: full *)
        END_IF;
    ELSIF local_deqEdge AND NOT local_enqEdge THEN
        IF local_count > 0 THEN
            (* Copy head element back to item. *)
            local_pSrc := local_pBufferBase;
            local_offset := local_head * local_elemSize;
            local_pSrc := local_pSrc + local_offset;
            local_pDst := local_pItemBase;
            local_copiedBytes := SysMemCpy(
                pbyDest := local_pDst,
                pbySource := local_pSrc,
                dwCount := TO_DWORD(local_elemSize)
            );

            local_head := (local_head + 1) MOD local_capacity;
            local_count := local_count - 1;
            status := 16#0000;
        ELSE
            status := 16#8001; (* dequeue rejected: empty *)
        END_IF;
    END_IF;
END_IF;

elementCount := local_count;
END_FUNCTION_BLOCK
